(* IEC 61131-3 sources: plc-vscode/tests/st/all/rusty/tests/lit/multi/polymorphism_fb, 5 files *)

(* ---- main.st ---- *)
FUNCTION main
    VAR
        instanceA: FbA;
        instanceB: FbB;
        instanceC: FbC;
        instanceD: FbD;

        refInstanceA: POINTER TO FbA;
    END_VAR

    refInstanceA := ADR(instanceA);
    refInstanceA^.alpha();
    refInstanceA^.bravo();
    refInstanceA^.charlie();
    refInstanceA^.delta();

    refInstanceA := ADR(instanceB);
    refInstanceA^.alpha();
    refInstanceA^.bravo();
    refInstanceA^.charlie();
    refInstanceA^.delta();

    refInstanceA := ADR(instanceC);
    refInstanceA^.alpha();
    refInstanceA^.bravo();
    refInstanceA^.charlie();
    refInstanceA^.delta();

    refInstanceA := ADR(instanceD);
    refInstanceA^.alpha();
    refInstanceA^.bravo();
    refInstanceA^.charlie();
    refInstanceA^.delta();
END_FUNCTION

(* ---- a.st ---- *)
FUNCTION_BLOCK FbA
    METHOD alpha
        printf('FbA::alpha$N');
    END_METHOD

    METHOD bravo
        printf('FbA::bravo$N');
    END_METHOD

    METHOD charlie
        printf('FbA::charlie$N');
    END_METHOD

    METHOD delta
        printf('FbA::delta$N');
    END_METHOD
END_FUNCTION_BLOCK

(* ---- b.st ---- *)
FUNCTION_BLOCK FbB EXTENDS FbA
    METHOD bravo
        printf('FbB::bravo$N');
    END_METHOD
END_FUNCTION_BLOCK

(* ---- c.st ---- *)
FUNCTION_BLOCK FbC EXTENDS FbB
    METHOD charlie
        printf('FbC::charlie$N');
    END_METHOD
END_FUNCTION_BLOCK

(* ---- d.st ---- *)
FUNCTION_BLOCK FbD EXTENDS FbC
    METHOD alpha
        printf('FbD::alpha$N');
    END_METHOD

    METHOD bravo
        printf('FbD::bravo$N');
    END_METHOD

    METHOD charlie
        printf('FbD::charlie$N');
    END_METHOD

    METHOD delta
        printf('FbD::delta$N');
    END_METHOD
END_FUNCTION_BLOCK
